{attribute 'qualified_only'}
{attribute 'strict'}
TYPE E_Error_Active_Module :
(
	noError := 0, Piston, Motor
);
END_TYPE

(* stored: Version 1.1.0.1, ProductVersion 3.1.4024.12
   DUT E_Error_Active_Module: Id {f52b7a91-0174-4891-bed2-fb6eec043efb} *)
